RoboDK station: PickPlace_Delta.rdk

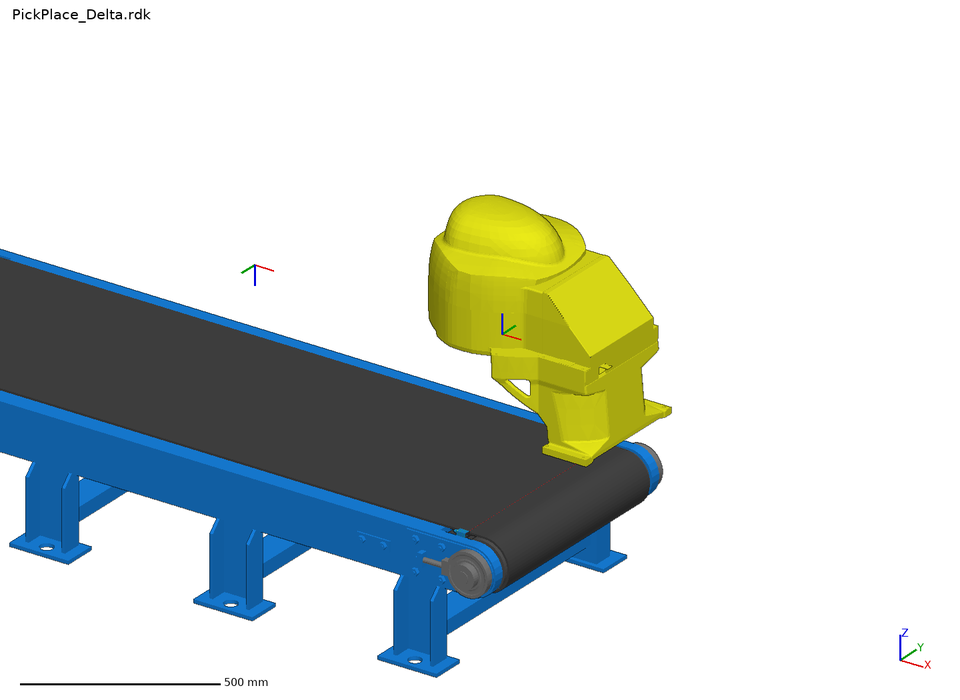
[picture v0: the station drawn from its stored meshes, robots at their saved joint values, targets as dots, program paths as lines]
Station PickPlace_Delta (saved by RoboDK 6.0.1). Poses are relative to the parent item; angles as X-Y-Z fixed-axis rotations.
Station parameters (name, value as stored): SICK WL4S Laser Sensor, 0
  - frame Conveyor Belt Wide (2m) Base at (0, 0, 0) mm
    - robot Conveyor Belt Wide (2m): 1 axes
        modified DH rows (alpha deg, a mm, theta deg, d mm): 0, 0, 0, 0 linear
        base shift (0, 0, 0) mm, rotated rx 0 ry 90 rz 0 deg
        joint limits [-900000] to [900000]; home [0]; saved at [-882707]
      - frame Conveyor Frame at (0, 0, 0) mm
        - object Box at (898881, 183.63, 2.38) mm, rotated rx -0.5 ry 0.33 rz 15.29 deg, size 50 x 100 x 25 mm, geometry from box.sld
        - object Box at (897722, 119.77, 3.01) mm, rotated rx -0.59 ry 0 rz -18.05 deg, size 50 x 100 x 25 mm, geometry from box.sld
        - object Box at (896441, 14.98, 4.04) mm, rotated rx -0.5 ry 0.32 rz 14.61 deg, size 50 x 100 x 25 mm, geometry from box.sld
        - object Box at (895254, 197, 2.25) mm, rotated rx -0.59 ry 0 rz -18.37 deg, size 50 x 100 x 25 mm, geometry from box.sld
    - frame Reference Box Frame at (60, 290, 366.5) mm
      - object ref_obj at (0, 0, 0) mm, size 252 x 305.4 x 216.7 mm, geometry from Box-12x10in-Closed.sld
      - object ref_lid at (-60, -186.65, 3.17) mm, rotated rx -0.56 ry 0.19 rz 0 deg, size 50 x 100 x 25 mm, geometry from box.sld
    - object SICK WL4S Laser Sensor at (1954, -20, 370) mm, rotated rx 180 ry 0 rz 90 deg, size 683.3 x 45.2 x 12.5 mm, geometry from SICK-WL4S-Laser-Sensor.sld
  - folder Python Scripts
    - Python program ConveyorReset (listed below)
    - Python program SensorReader (listed below)
    - Python program ConveyorRunner (listed below)
    - Python program BoxSpawner (listed below)
  - program MainProgram (5 instructions, listed below)
  - notes Description: <!DOCTYPE HTML PUBLIC "-//W3C//DTD HTML 4.0//EN" "http://www.w3.org/TR/REC-html40/strict.dtd">
<html><head><meta name="qrichtext" content="1" /><style type="text/css">
p, li { white-space: pre-wrap; }
</style></head><body style=" font-family:'MS Shell Dlg 2'; font-size:8.25pt; font-weight:400; font-style:normal;">
<p style=" margin-top:0px; margin-bottom:0px; margin-left:0px; margin-right:0px; -qt-block-indent:0; text-indent:0px;">This example demonstrates a conveyor simulation in RoboDK using Python scripting. A script generates boxes of varying sizes and positions while the conveyor moves continuously. A sensor detects when a box reaches the conveyor’s edge and stops the conveyor. The station showcases how conveyors, part generation, and sensor-based control can be simulated with the API.</p></body></html>
  - frame Fanuc M-1iA/0.5SL Base at (1954.3, 143.51, 858.22) mm
    - robot Fanuc M-1iA/0.5SL: 4 axes, payload 0.5 kg, reach 420 mm, repeatability 0.03 mm, weight 23 kg
        joint limits [-25, -25, -25, -36000] to [80, 80, 80, 36000]; home [0, 0, 0, 0]; saved at [65.567, 65.567, 65.567, 0]
      - tool Tool 1, TCP at (0, 0, 0) mm
  - frame CamFrame at (1207.08, 136.9, 843.5) mm, rotated rx -180 ry -0.2 rz -0.44 deg
    - camera Camera 1
  - frame Frame 6 at (5.31, 161.47, 358.87) mm, rotated rx 0 ry 0 rz 90 deg

--- Python program ConveyorReset ---
# Type help("robodk.robolink") or help("robodk.robomath") for more information
# Press F5 to run the script
# Documentation: https://robodk.com/doc/en/RoboDK-API.html
# Reference:     https://robodk.com/doc/en/PythonAPI/robodk.html
# Note: It is not required to keep a copy of this file, your Python script is saved with your RDK project

from robodk import robolink  # RoboDK API
from robodk import robomath  # Robot toolbox

#---------------------------------------
# Avoid auto-select
RDK = robolink.Robolink()
RDK.setSelection([])

#---------------------------------------
# Get the conveyor
conveyors = [x for x in RDK.ItemList(robolink.ITEM_TYPE_ROBOT_AXES) if len(x.Joints().tolist()) == 1 and 'conveyor' in x.Name().lower()]
if not conveyors:
    RDK.ShowMessage('No conveyor found. Please add a conveyor with "conveyor" in its name, i.e. "Conveyor Belt"')
    quit()
conveyor = RDK.ItemUserPick(itemtype_or_list=conveyors) if len(conveyors) > 1 else conveyors[0]
if not conveyor.Valid():
    quit()
print(f'Using conveyor: {conveyor.Name()}')
conveyor_min, conveyor_max, _ = conveyor.JointLimits()

#---------------------------------------
# Get the conveyor's reference frame
frames = [x for x in conveyor.Childs() if x.Type() == robolink.ITEM_TYPE_FRAME]
if not frames:
    frames = [RDK.AddFrame(conveyor.Name() + ' Frame', conveyor)]
conveyor_frame = RDK.ItemUserPick(itemtype_or_list=frames) if len(frames) > 1 else frames[0]
if not conveyor_frame.Valid():
    quit()
print(f'Using conveyor frame: {conveyor_frame.Name()}')
conveyor_frame.setVisible(False)
conveyor_frame.setParam("Tree", "Collapse")

#---------------------------------------
# Reset the conveyor
RDK.Render(False)
for child in conveyor_frame.Childs():
    if child.Type() == robolink.ITEM_TYPE_OBJECT and 'box' in child.Name().lower():
        child.Delete()
conveyor.setJoints(conveyor_min)
RDK.Render(True)

--- Python program SensorReader ---
# Type help("robodk.robolink") or help("robodk.robomath") for more information
# Press F5 to run the script
# Documentation: https://robodk.com/doc/en/RoboDK-API.html
# Reference:     https://robodk.com/doc/en/PythonAPI/robodk.html
# Note: It is not required to keep a copy of this file, your Python script is saved with your RDK project

from robodk import robolink  # RoboDK API
from robodk import robomath  # Robot toolbox
import time

#---------------------------------------
# Settings

# Prefer the Sensor plugin, as it is much more reliable!
# More info here: https://github.com/RoboDK/Plug-In-Interface/tree/master/PluginCollisionSensor
USE_SENSOR_PLUGIN = True
SENSOR_PLUGIN_DLL = 'PluginCollisionSensor.dll'
SENSOR_PLUGIN_NAME = 'Plugin Collision Sensor'

#---------------------------------------
# Enable the sensor plugin
RDK = robolink.Robolink()
RDK.setSelection([])  # Avoid auto-select with ItemUserPick

if USE_SENSOR_PLUGIN:
    status = RDK.Command('PluginLoad', SENSOR_PLUGIN_DLL)
    if status != 'OK':
        RDK.ShowMessage(f'Sensor: Using Python script (failed to load {SENSOR_PLUGIN_NAME})', False)
        USE_SENSOR_PLUGIN = False

#---------------------------------------
# Get the sensor item
sensors = [x for x in RDK.ItemList(robolink.ITEM_TYPE_OBJECT) if 'sensor' in x.Name().lower()]
if not sensors:
    RDK.ShowMessage('No sensor found. Please add a sensor object with "sensor" in its name, i.e. "Laser Sensor"')
    quit()
sensor = RDK.ItemUserPick(itemtype_or_list=sensors) if len(sensors) > 1 else sensors[0]
if not sensor.Valid():
    quit()
SENSOR_IO = sensor.Name()
print(f'Using laser sensor: {SENSOR_IO}')

#---------------------------------------
# Enable the sensor item
if USE_SENSOR_PLUGIN:
    status = RDK.PluginCommand(SENSOR_PLUGIN_NAME, "Activate", SENSOR_IO)
    if 'OK' == status:
        RDK.ShowMessage(f'Sensor: Using {SENSOR_PLUGIN_NAME}', False)
        quit()

RDK.ShowMessage('Sensor: Using Python script', False)
USE_SENSOR_PLUGIN = False

#---------------------------------------
# Get the conveyor
conveyors = [x for x in RDK.ItemList(robolink.ITEM_TYPE_ROBOT_AXES) if len(x.Joints().tolist()) == 1 and 'conveyor' in x.Name().lower()]
if not conveyors:
    RDK.ShowMessage('No conveyor found. Please add a conveyor with "conveyor" in its name, i.e. "Conveyor Belt"')
    quit()
conveyor = RDK.ItemUserPick(itemtype_or_list=conveyors) if len(conveyors) > 1 else conveyors[0]
if not conveyor.Valid():
    quit()
print(f'Using conveyor: {conveyor.Name()}')

#---------------------------------------
# Get the conveyor's reference frame
frames = [x for x in conveyor.Childs() if x.Type() == robolink.ITEM_TYPE_FRAME]
if not frames:
    frames = [RDK.AddFrame(conveyor.Name() + ' Frame', conveyor)]
conveyor_frame = RDK.ItemUserPick(itemtype_or_list=frames) if len(frames) > 1 else frames[0]
if not conveyor_frame.Valid():
    quit()
print(f'Using conveyor frame: {conveyor_frame.Name()}')

while True:

    time.sleep(0.01)

    detection = 0
    childs = conveyor_frame.Childs()
    for box in [x for x in childs if x.Type() == robolink.ITEM_TYPE_OBJECT]:
        if box.Valid(True) and RDK.Collision(sensor, box):
            detection = 1
            break

    RDK.setParam(SENSOR_IO, detection)

--- Python program ConveyorRunner ---
# Type help("robodk.robolink") or help("robodk.robomath") for more information
# Press F5 to run the script
# Documentation: https://robodk.com/doc/en/RoboDK-API.html
# Reference:     https://robodk.com/doc/en/PythonAPI/robodk.html
# Note: It is not required to keep a copy of this file, your Python script is saved with your RDK project

from robodk import robolink  # RoboDK API
from robodk import robomath  # Robot toolbox
import time

#---------------------------------------
# Avoid auto-select
RDK = robolink.Robolink()
RDK.setSelection([])

#---------------------------------------
# Get the sensor
sensors = [x for x in RDK.ItemList(robolink.ITEM_TYPE_OBJECT) if 'sensor' in x.Name().lower()]
if not sensors:
    RDK.ShowMessage('No sensor found. Please add a sensor object with "sensor" in its name, i.e. "Laser Sensor"')
    quit()
sensor = RDK.ItemUserPick(itemtype_or_list=sensors) if len(sensors) > 1 else sensors[0]
if not sensor.Valid():
    quit()
SENSOR_IO = sensor.Name()
print(f'Using laser sensor: {SENSOR_IO}')

#---------------------------------------
# Get the conveyor
conveyors = [x for x in RDK.ItemList(robolink.ITEM_TYPE_ROBOT_AXES) if len(x.Joints().tolist()) == 1 and 'conveyor' in x.Name().lower()]
if not conveyors:
    RDK.ShowMessage('No conveyor found. Please add a conveyor with "conveyor" in its name, i.e. "Conveyor Belt"')
    quit()
conveyor = RDK.ItemUserPick(itemtype_or_list=conveyors) if len(conveyors) > 1 else conveyors[0]
if not conveyor.Valid():
    quit()
print(f'Using conveyor: {conveyor.Name()}')
conveyor_min, conveyor_max, _ = conveyor.JointLimits()
conveyor_max = conveyor_max.list()[0]

while True:

    time.sleep(0.01)

    sensor_state = RDK.getParam(SENSOR_IO)
    if sensor_state == 1:
        conveyor.Stop()
    elif not conveyor.Busy():
        target = [min(conveyor_max, conveyor.Joints().list()[0] + 99999)]  # this is to avoid lengthy calculations when the target is to far away (as oppose to conveyor.MoveJ(conveyor_max, False))
        conveyor.MoveJ(target, False)

--- Python program BoxSpawner ---
# Type help("robodk.robolink") or help("robodk.robomath") for more information
# Press F5 to run the script
# Documentation: https://robodk.com/doc/en/RoboDK-API.html
# Reference:     https://robodk.com/doc/en/PythonAPI/robodk.html
# Note: It is not required to keep a copy of this file, your Python script is saved with your RDK project

from robodk import robolink  # RoboDK API
from robodk import robomath  # Robot toolbox
import time
import random

RANDOMIZE_SIZE = True
SIZE_RANGE_FACTOR = [0.5, 0.9]  # %/100, minimum and maximum scale

RANDOMIZE_ROTATION = True
ROTATION_MAX = 20  # degrees, maximum rotation along reference Z (+/-)

RANDOMIZE_POSITION = True
POSITION_MAX = 100  # mm, maximum lateral offset (+/-)

#---------------------------------------
# Avoid auto-select
RDK = robolink.Robolink()
RDK.setSelection([])

#---------------------------------------
# Get the reference box
boxes = [x for x in RDK.ItemList(robolink.ITEM_TYPE_OBJECT) if 'box' in x.Name().lower() and 'ref' in x.Name().lower()]
if not boxes:
    RDK.ShowMessage('No reference box found. Please add a reference box with "box" and "ref" in its name, i.e. "Reference Box"')
    quit()
ref_box = RDK.ItemUserPick(itemtype_or_list=boxes) if len(boxes) > 1 else boxes[0]
if not ref_box.Valid():
    quit()
print(f'Using reference box: {ref_box.Name()}')
ref_box.setVisible(False)
ref_box.Parent().setParam('Tree', 'Collapse')

#---------------------------------------
# Get the conveyor
conveyors = [x for x in RDK.ItemList(robolink.ITEM_TYPE_ROBOT_AXES) if len(x.Joints().tolist()) == 1 and 'conveyor' in x.Name().lower()]
if not conveyors:
    RDK.ShowMessage('No conveyor found. Please add a conveyor with "conveyor" in its name, i.e. "Conveyor Belt"')
    quit()
conveyor = RDK.ItemUserPick(itemtype_or_list=conveyors) if len(conveyors) > 1 else conveyors[0]
if not conveyor.Valid():
    quit()
print(f'Using conveyor: {conveyor.Name()}')

#---------------------------------------
# Get the conveyor's reference frame
frames = [x for x in conveyor.Childs() if x.Type() == robolink.ITEM_TYPE_FRAME]
if not frames:
    frames = [RDK.AddFrame(conveyor.Name() + ' Frame', conveyor)]
conveyor_frame = RDK.ItemUserPick(itemtype_or_list=frames) if len(frames) > 1 else frames[0]
if not conveyor_frame.Valid():
    quit()
print(f'Using conveyor frame: {conveyor_frame.Name()}')


def spawn_box():
    # Copy/paste changes the user selection
    RDK.Render(False)
    selection = RDK.Selection()
    ref_box.Copy(copy_children=False)
    new_box = ref_box.Parent().Paste()
    RDK.setSelection(selection)
    new_box.setVisible(False)
    new_box.setName('Box')

    pose = new_box.Pose()
    if RANDOMIZE_SIZE:
        scale = random.uniform(SIZE_RANGE_FACTOR[0], SIZE_RANGE_FACTOR[1])
        new_box.Scale(scale)

    if RANDOMIZE_POSITION:
        lateral_offset = random.uniform(-POSITION_MAX, POSITION_MAX)  # Assuming reference frame has Y crossing the conveyor's width
        pose = robomath.RelTool(pose, 0, lateral_offset, 0)

    if RANDOMIZE_ROTATION:
        rotation = random.uniform(-ROTATION_MAX, ROTATION_MAX)
        pose = robomath.RelTool(pose, 0, 0, 0, 0, 0, rotation)

    new_box.setPose(pose)
    RDK.Render(False)  # Update pose

    new_box.setParentStatic(conveyor_frame)
    new_box.setVisible(True)
    RDK.Render(True)
    return new_box


box_queue = conveyor_frame.Childs()
while True:

    time.sleep(0.1)

    # Remove boxes removed from the conveyor, deleted or too far away
    childs = conveyor_frame.Childs()
    for box in box_queue:
        if not box.Valid(True) or box not in childs:
            box_queue.remove(box)

    if not box_queue:
        box_queue.append(spawn_box())
        continue

    # Spawn new boxes if space is sufficient
    if box_queue[-1].Valid(True) and not RDK.Collision(ref_box, box_queue[-1]):
        box_queue.append(spawn_box())

--- program MainProgram (robot Conveyor Belt Wide (2m)) ---
  Call ConveyorReset
  Run SensorReader
  Set speed (25.0 mm/s)
  Run ConveyorRunner
  Run BoxSpawner
